TYPE E_2OO3_MODE :
(
    MODE_2OO3 := 0,
    IG1 := 1,
    IG2 := 2,
    IG3 := 3
);
END_TYPE

(* stored: Version 1.1.0.1
   DUT E_2OO3_MODE: Id {7da80cf0-4fde-4ce3-82c4-7c1c74badc27} *)
